TYPE "ST_DeclarationOutCmd"
VERSION : 0.1
   STRUCT
      "Result" : DInt;
   END_STRUCT;
END_TYPE
